FUNCTION_BLOCK NFHDiag (* Basic Function Block Type *)
  (* Standard: 61499-2 *)
  (* Version 0.0, 10/6/2026, Schneider Electric, Template *)
  PACKAGE SE.Nereda;
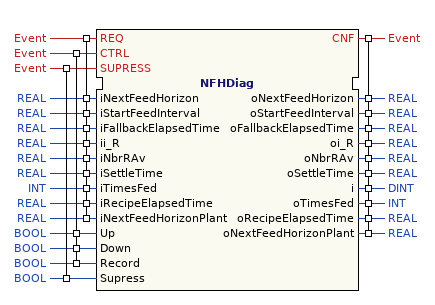
  EVENT_INPUT
    REQ WITH iNextFeedHorizon, iStartFeedInterval, iFallbackElapsedTime, ii_R, iSettleTime, iNbrRAv, iTimesFed, iRecipeElapsedTime, iNextFeedHorizonPlant; (* Normal Execution Request *)
    CTRL WITH Up, Down, Record;
    SUPRESS WITH Supress;
  END_EVENT
  EVENT_OUTPUT
    CNF WITH oNextFeedHorizon, oStartFeedInterval, oFallbackElapsedTime, oi_R, oSettleTime, i, oNbrRAv, oTimesFed, oRecipeElapsedTime, oNextFeedHorizonPlant; (* Execution Confirmation *)
  END_EVENT
  VAR_INPUT
    iNextFeedHorizon : REAL;
    iStartFeedInterval : REAL;
    iFallbackElapsedTime : REAL;
    ii_R : REAL;
    iNbrRAv : REAL;
    iSettleTime : REAL;
    iTimesFed : INT;
    iRecipeElapsedTime : REAL;
    iNextFeedHorizonPlant : REAL;
    Up : BOOL;
    Down : BOOL;
    Record : BOOL;
    Supress : BOOL;
  END_VAR
  VAR_OUTPUT
    oNextFeedHorizon : REAL;
    oStartFeedInterval : REAL;
    oFallbackElapsedTime : REAL;
    oi_R : REAL;
    oNbrRAv : REAL;
    oSettleTime : REAL;
    i : DINT;
    oTimesFed : INT;
    oRecipeElapsedTime : REAL;
    oNextFeedHorizonPlant : REAL;
  END_VAR
  VAR
    NextFeedHorizon : ARRAY [0..99] OF REAL;
    StartFeedInterval : ARRAY [0..99] OF REAL;
    FallbackElapsedTime : ARRAY [0..99] OF REAL;
    NbrRAv : ARRAY [0..99] OF REAL;
    i_R : ARRAY [0..99] OF REAL;
    SettleTime : ARRAY [0..99] OF REAL;
    TimesFed : ARRAY [0..99] OF INT;
    RecipeElapsedTime : ARRAY [0..99] OF REAL;
    NextFeedHorizonPlant : ARRAY [0..99] OF REAL;
  END_VAR
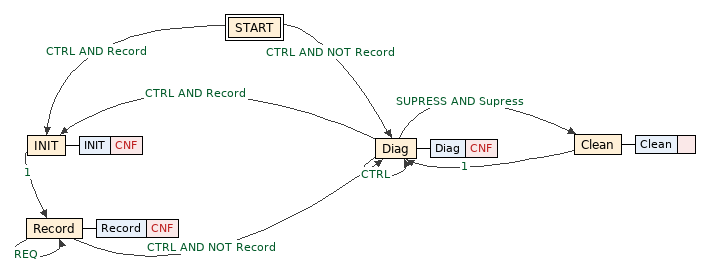
  EC_STATES
    START; (* Initial State *)
    Record : Record -> CNF;
    Diag : Diag -> CNF;
    INIT : INIT -> CNF;
    Clean : Clean;
  END_STATES
  EC_TRANSITIONS
    START TO INIT := CTRL AND Record;
    START TO Diag := CTRL AND NOT Record;
    Diag TO INIT := CTRL AND Record;
    Record TO Record := REQ;
    Diag TO Diag := CTRL;
    Record TO Diag := CTRL AND NOT Record;
    INIT TO Record := 1;
    Diag TO Clean := SUPRESS AND Supress;
    Clean TO Diag := 1;
  END_TRANSITIONS
  ALGORITHM Record IN ST:
;
IF i < 100 THEN
	NextFeedHorizon[i] := iNextFeedHorizon;
	StartFeedInterval[i] := iStartFeedInterval;
	FallbackElapsedTime[i] := iFallbackElapsedTime;
	NbrRAv[i] := iNbrRAv;
	i_R[i] := ii_R;
	SettleTime[i] := iSettleTime;
	TimesFed[i] := iTimesFed;
	RecipeElapsedTime[i] := iRecipeElapsedTime;
	NextFeedHorizonPlant[i] := iNextFeedHorizonPlant;

	i := i + 1;
END_IF;

REQ := FALSE;
  END_ALGORITHM
  ALGORITHM Diag IN ST:
;
IF Up AND NOT Down THEN
	i := i + 1;
ELSIF NOT Up AND Down THEN
	i := i - 1;
END_IF;

oNextFeedHorizon := NextFeedHorizon[i];
oStartFeedInterval := StartFeedInterval[i];
oFallbackElapsedTime := FallbackElapsedTime[i];
oNbrRAv := NbrRAv[i];
oi_R := i_R[i];
oSettleTime := SettleTime[i];
oTimesFed := TimesFed[i];
oRecipeElapsedTime := RecipeElapsedTime[i];
oNextFeedHorizonPlant := NextFeedHorizonPlant[i];

CTRL := FALSE;
  END_ALGORITHM
  ALGORITHM INIT IN ST:
;
i := 0;
  END_ALGORITHM
  ALGORITHM Clean IN ST:
;
FOR i := 0 TO 98 DO
	NextFeedHorizon[i] := 0;
	StartFeedInterval[i] := 0;
	FallbackElapsedTime[i] := 0;
	NbrRAv[i] := 0;
	i_R[i] := 0;
	SettleTime[i] := 0;
	TimesFed[i] := 0;
	RecipeElapsedTime[i] := 0;
	NextFeedHorizonPlant[i] := 0;
END_FOR;
  END_ALGORITHM
END_FUNCTION_BLOCK
